(*
	Contract for span processors. FB_TracerProvider stages processors each scan, then its tick
	passes every ended span to onEnd of each staged processor and releases the span once they
	have all returned. The span is borrowed: a processor that keeps it past onEnd must clone it.
*)
FUNCTION_BLOCK ABSTRACT FB_SpanProcessor_Base

(* Extension point that may change the span before it is exported. *)
METHOD ABSTRACT enrich
VAR_IN_OUT
	span: FB_Span;
END_VAR
END_METHOD

METHOD ABSTRACT free
END_METHOD

(* Called once for each ended span. The span is borrowed and released after the call. *)
METHOD ABSTRACT onEnd
VAR_INPUT
	span: REFERENCE TO FB_Span;
END_VAR
END_METHOD

PROPERTY pSelf : POINTER TO FB_SpanProcessor_Base
GET
pSelf := THIS;
END_GET
END_PROPERTY

(* Called once per provider tick, after the ended spans have been handed out. *)
METHOD ABSTRACT tick
END_METHOD

END_FUNCTION_BLOCK

(* stored: Version 1.1.0.1
   POU FB_SpanProcessor_Base: Id {59b7378e-f835-4bd4-a5bd-0e08f64b62dc}, SpecialFunc None
   Method enrich: Id {82915b2d-b9e0-488c-b46c-2bddccb07065}
   Method free: Id {8921e54d-7ee7-4ebc-b99f-15368644b974}
   Method onEnd: Id {7d1578d8-6be9-45c4-8a55-2d5219356e6c}
   Property pSelf: Id {747c4406-fcd5-441e-9545-c175f6a7aad9}
   Get Get: Id {50e07d9a-e8c7-4fdb-9304-e250405b4795}
   Method tick: Id {ab265dbc-fe04-402c-a2ab-a835cd7e80e6} *)
